// TIA Portal V19 export
TYPE "ST_Pos"
   STRUCT
      X : Int;
      Y : Int;
      Z : Int;
      Rz : Int;
      Valid : Bool;
   END_STRUCT;
END_TYPE
